(* IEC 61131-3 sources: s22-soft-shell/st_interpret/tests/test_inputs/misc, 5 files *)

(* ---- intidentityfunction.st ---- *)
FUNCTION IntIdentityFunction : INT

VAR_INPUT
  Input1 :	INT;
END_VAR

  IntIdentityFunction := Input1;
END_FUNCTION

(* ---- nestedaddfunction.st ---- *)
FUNCTION NestedAddFunction : INT //INT is the return parameter data type
VAR_INPUT
  Input1 :	INT; //Input parameter 1 to the function
  Input2 :	INT; //Input parameter 2 to the function
END_VAR

VAR
  Sum :	INT; //Local variable for temporary calculation
END_VAR

  Sum := IntIdentityFunction(Input1) + Input2; //Total sum

  NestedAddFunction := Sum; //Set the return parameter

END_FUNCTION

(* ---- simpleaddfunction.st ---- *)
FUNCTION SimpleAddFunction : INT //INT is the return parameter data type
VAR_INPUT
  Input1 :	INT; //Input parameter 1 to the function
  Input2 :	INT; //Input parameter 2 to the function
END_VAR

VAR
  Sum :	INT; //Local variable for temporary calculation
END_VAR

  Sum:= Input1 + Input2; //Total sum

  SimpleAddFunction:= Sum; //Set the return parameter

END_FUNCTION

(* ---- 09_Main_Add.st ---- *)
//Testing simple function call to add two numbers together
PROGRAM 09_Main_Add
    VAR
	a : int;
        b : int;
        result0 : int;
        result1 : int;
        result2 : int;
        result3 : int;
    END_VAR
        a := 3;
        b := 5;

        // four different ways of function input
        result0 := SimpleAddFunction(10, 10+5); // expects outputs of 25

        result1 := SimpleAddFunction(Input1 := 5, Input2 := 10); // expects outputs of 15

        result2 := SimpleAddFunction(a, b); // expects outputs of 8

        result3 := SimpleAddFunction(Input1 := a, Input2 := b); // expects outputs of 8

END_PROGRAM

(* ---- 09_Main_Add_Nested.st ---- *)
// Function call to add two numbers together, which itself contains another function call
PROGRAM 09_Main_Add
    VAR
	a : int;
        b : int;
        result0 : int;
        result1 : int;
        result2 : int;
        result3 : int;
    END_VAR
        a := 3;
        b := 5;

        // four different ways of function input
        result0 := NestedAddFunction(10, 10+5); // expects outputs of 25

        result1 := NestedAddFunction(Input1 := 5, Input2 := 10); // expects outputs of 15

        result2 := NestedAddFunction(a, b); // expects outputs of 8

        result3 := NestedAddFunction(Input1 := a, Input2 := b); // expects outputs of 8

END_PROGRAM
